Fanuc KAREL source: kd00048.KL

PROGRAM KD00048
%STACKSIZE=65535
%PRIORITY=65535
%NOLOCKGROUP
VAR
I : INTEGER
J : INTEGER
B : BOOLEAN
R : REAL
S : STRING[80]
-- UNRESOLVED DECLARATIONS (source type spelling not recovered)
-- PTH : TYPE_0x001F (type_u16=0x001F)
BEGIN
-- UNRESOLVED_PC line 12 opcodes [01 22 1C 9D 2C 08 82 0B] marker_code=0
END KD00048
